(* IEC 61131-3 sources: ISA-88-Bioreactor-Automation-Template-DE-IE/ISA-88-Bioreactor-Automation-Template-DE-IE.fbsdev/ThermalManager.iecapp^/FunctionBlocks, 4 files *)

(* ---- ThermalAlarm_FB_ST.fb.st ---- *)
FUNCTION_BLOCK ThermalAlarm_FB_ST
VAR_INPUT
    Tn_Temp_Value : REAL;   // current tank temperature
    Tn_Temp_Max   : REAL;   // maximum safe temperature
END_VAR

VAR_OUTPUT
    Thermal_Alarm : BOOL := FALSE;
END_VAR

// Alarm logic
IF Tn_Temp_Value > Tn_Temp_Max THEN
    Thermal_Alarm := TRUE;
ELSE
    Thermal_Alarm := FALSE;
END_IF;

(* ---- ThermalControl_FB_ST.fb.st ---- *)
FUNCTION_BLOCK ThermalControl_FB_ST
VAR_INPUT
    Cycle_Active     : BOOL;   // cycle running
    Mix_Complete     : BOOL;   // mixing finished
    Tn_Temp_Value    : REAL;   // current temperature
    Tn_Temp_Setpoint : REAL;   // desired setpoint
END_VAR

VAR_OUTPUT
    Heater           : BOOL := FALSE;
    Heat_Complete    : BOOL := FALSE;
END_VAR

// Heat control logic
IF Cycle_Active AND Mix_Complete THEN
    Heater := (Tn_Temp_Value < Tn_Temp_Setpoint);
    IF Tn_Temp_Value >= Tn_Temp_Setpoint THEN
        Heat_Complete := TRUE;
        Heater := FALSE;
    END_IF;
ELSE
    Heater := FALSE;
    Heat_Complete := FALSE;
END_IF;

(* ---- ThermalInterlock_FB_ST.fb.st ---- *)
FUNCTION_BLOCK ThermalInterlock_FB_ST
VAR_INPUT
    Pump_Discharge : BOOL; // pump running
    Mixer_Motor    : BOOL; // mixer running
END_VAR

VAR_OUTPUT
    Thermal_Enable : BOOL := FALSE;
END_VAR

// Interlock logic
Thermal_Enable := NOT (Pump_Discharge OR Mixer_Motor);

(* ---- ThermalTimer_FB_ST.fb.st ---- *)
FUNCTION_BLOCK ThermalTimer_FB_ST
VAR_INPUT
    Cycle_Active : BOOL;   // overall cycle running
    Mix_Complete : BOOL;   // mixing finished
    PT           : TIME := T#15s; // preset Thermaling time (adjust as needed)
END_VAR

VAR_OUTPUT
    ThermalTimer_Done : BOOL := FALSE;
END_VAR

VAR
    TON_Thermal : TON; // IEC timer instance
END_VAR

// Timer logic
TON_Thermal(IN := (Cycle_Active AND Mix_Complete), PT := PT);

ThermalTimer_Done := TON_Thermal.Q;
